(* IEC 61131-3 sources: codesys-to-s7/tests/corpus/C2S7-NAME-KEYWORD/pos, 1 file *)

(* ---- input.st ---- *)
FUNCTION_BLOCK FB_Case
VAR
    begin : INT;
END_VAR
begin := 1;
END_FUNCTION_BLOCK
